// TIA Portal V20 export
// export: Created 2026-10-20T12:46:53.1203727Z, ExportSetting WithDefaults, DisplayName Totally Integrated Automation Portal, DisplayVersion V20 Update 6, DisplayName TIA Portal Openness, DisplayVersion V20 Update 6, DisplayName TIA Portal Version Control Interface, DisplayVersion V20 Update 6, DisplayName SINAMICS Startdrive Advanced, DisplayVersion V20 SP1, DisplayName SINAMICS Startdrive G130, G150, S120, S150, SINAMICS MV, G220, S200, S210, DisplayVersion V20 SP1, DisplayName SINAMICS Startdrive G110M, G120, G120C, G120D, G120P, G115D, DisplayVersion V20 SP1, DisplayName STEP 7 Professional, DisplayVersion V20 Update 6, DisplayName STEP 7 Safety, DisplayVersion V20 Update 2, DisplayName WinCC Basic/Comfort/Advanced, DisplayVersion V20 Update 6, DisplayName WinCC Unified, DisplayVersion V20 Update 6
FUNCTION "ParseShuttle_Status" : "Shuttle_MQTT_Status_Msg"   // FC16, SCL
{ S7_Optimized_Access := 'TRUE' }
VERSION : 0.1
// stored: AutoNumber true, IsIECCheckEnabled false, SetENOAutomatically false, UDAEnableTagReadback false
   VAR_INPUT
      String_1 : String;
      String_2 : String;
      String_3 : String;
      String_4 : String;
      String_5 : String;
      String_6 : String;
   END_VAR
   VAR CONSTANT
      Empty : String;
   END_VAR
BEGIN
   #ParseShuttle_Status.Request_ID := "FindDINTFieldFragmented"(FieldName := 'requestId',
                                                                Str1 := #String_1,
                                                                Str2:=#Empty);
   #ParseShuttle_Status.Position_ID := "FindDINTFieldFragmented"(FieldName := 'positionId',
                                                                 Str1 := #String_1,
                                                                 Str2 := #Empty);
   #ParseShuttle_Status.Destination_ID := "FindDINTFieldFragmented"(FieldName := 'destinationId',
                                                                    Str1 := #String_1,
                                                                    Str2:=#Empty);
   #ParseShuttle_Status.Distance_Remaining := "FindDINTFieldFragmented"(FieldName := 'distanceRemaining',
                                                                        Str1 := #String_1,
                                                                        Str2 := #Empty);
   #ParseShuttle_Status.Position_X := "FindDINTFieldFragmented"(FieldName := 'positionX',
                                                                Str1 := #String_1,
                                                                Str2 := #Empty);
   #ParseShuttle_Status.Position_Y := "FindDINTFieldFragmented"(FieldName := 'positionY',
                                                                Str1 := #String_1,
                                                                Str2 := #Empty);
   #ParseShuttle_Status.Floor := "FindIntField"(FieldName := 'floor',
                                                   JsonStr := #String_1);
   #ParseShuttle_Status.Operation_Mode := "FindStringField"(FieldName := 'operationMode',
                                                            JsonStr := #String_1);
   #ParseShuttle_Status.Operational_State := "FindStringField"(FieldName := 'operationState',
                                                               JsonStr := #String_2);
   #ParseShuttle_Status.Load_State := "FindStringField"(FieldName := 'loadState',
                                                        JsonStr := #String_2);
   #ParseShuttle_Status.Error_Vehicle_1 := INT_TO_UINT("FindINTFieldFragmented"(FieldName := 'errorVehicle1',
                                                                                                                                    Str1 := #String_2,
                                                                                                                                    Str2:=#String_2));
   #ParseShuttle_Status.Error_Vehicle_2 := INT_TO_UINT("FindIntField"(FieldName := 'errorVehicle2',
                                                                                                                          JsonStr := #String_2));
   #ParseShuttle_Status.Error_Vehicle_3 := INT_TO_UINT("FindIntField"(FieldName := 'errorVehicle3',
                                                                                                                          JsonStr := #String_3));
   #ParseShuttle_Status.Error_Vehicle_4 := INT_TO_UINT("FindIntField"(FieldName := 'errorVehicle4',
                                                                                                                          JsonStr := #String_3));
   #ParseShuttle_Status.Error_Vehicle_5 := INT_TO_UINT("FindIntField"(FieldName := 'errorVehicle5',
                                                                                                                          JsonStr := #String_3));
   #ParseShuttle_Status.Error_Vehicle_6 := INT_TO_UINT("FindIntField"(FieldName := 'errorVehicle6',
                                                                                                                          JsonStr := #String_4));
   #ParseShuttle_Status.Sensor_Inputs := INT_TO_UINT("FindIntField"(FieldName := 'sensorInputs',
                                                                                                                      JsonStr := #String_4));
   #ParseShuttle_Status.Sensor_Outputs := INT_TO_UINT("FindIntField"(FieldName := 'sensorOutputs',
                                                                                                                        JsonStr := #String_4));
   #ParseShuttle_Status.Reader_Value := "FindDINTFieldFragmented"(FieldName := 'readerValue',
                                                                  Str1 := #String_4,
                                                                Str2 := #Empty);
   #ParseShuttle_Status.Pallet_Type := "FindStringField"(FieldName := 'palletType',
                                                         JsonStr := #String_4);
   #ParseShuttle_Status.Energy_Level := INT_TO_UINT("FindINTFieldFragmented"(FieldName := 'energyLevel',
                                                                                                                              Str1 := #String_5,
                                                                                                                              Str2:=#String_5));
   #ParseShuttle_Status.Battery_Voltage := INT_TO_UINT("FindIntField"(FieldName := 'batteryVoltage',
                                                                                                                          JsonStr := #String_5));
   #ParseShuttle_Status.Paused := "FindBoolField"(FieldName := 'paused',
                                                  JsonStr := #String_5);
   #ParseShuttle_Status.Last_Received_Order_ID := "FindIntField"(FieldName := 'lastReceivedOrderId',
                                                                 JsonStr := #String_5);
    #ParseShuttle_Status.Current_Order_ID := "FindIntField"(FieldName := 'currentOrderId',
                                                            JsonStr := #String_6);
          #ParseShuttle_Status.Last_Finished_Order_ID := "FindIntField"(FieldName := 'lastFinishedOrderId',
                                                                        JsonStr := #String_6);
END_FUNCTION
